(* CODESYS project PLC Pool Water Level Control Program.export

Project tree, tasks and I/O mapping:
  Device : CODESYS Control Win V3 x64, CODESYS, version 3.5.22.40
    application Application
      libraries: Standard, 3.5.22.0 (System)
      task MainTask (cyclic, interval t#100ms, priority 1) calls PLC_PRG [Read level and calculate pump command], TankSimulation [Use the command to calculate the new tank volume], TrialTester, TuningManager
      task VISU_TASK (cyclic, interval 100 ms, priority 31) calls VisuElems.Visu_Prg
      program PLC_PRG [LD]
      function block PoolModel [ST]
      program TankSimulation [ST]
      program TrialTester [ST]
      program TuningManager [ST]
      function block TuningTrial [ST]
      function block Twiddle [ST]
      function block ValveController [ST]
      visualisation TankOverview
*)

// Device/Application/PLC_PRG
PROGRAM PLC_PRG
VAR
	AutomationEnabled: BOOL; // FALSE means system is in manual mode
	ValveCommand : REAL := 0.0; // this is the precent-open that the valve needs to be
	FillingRequest : BOOL := FALSE;
	LowLevel : BOOL := FALSE; // when tank reaches 30% or less
	HighLevel : BOOL := FALSE; // when tank reaches 80% or more
	Trip : BOOL := FALSE; // activated automatically when HighHigh becomes TRUE
	ResetTrip : BOOL := FALSE;  // activated by operator switch
	
	// configure the controller
	LevelController : ValveController;
END_VAR

VAR_INPUT
	PoolLevelDeviation : REAL := 0.0; // inches
	HighHigh : BOOL := FALSE; // when level reaches 95% due to a system errors
	ActiveKp : REAL := 40.0;
	ActiveKi : REAL := 1.0;
END_VAR

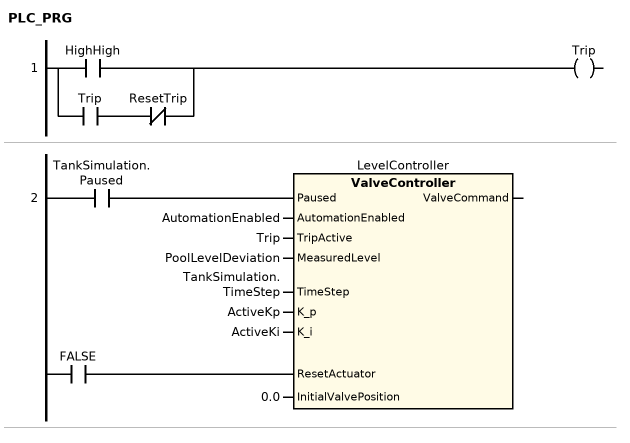
// NETWORK 1
Trip := HighHigh OR Trip AND NOT ResetTrip;

// NETWORK 2
LevelController(
    Paused := TankSimulation.Paused,
    AutomationEnabled := AutomationEnabled,
    TripActive := Trip,
    MeasuredLevel := PoolLevelDeviation,
    TimeStep := TankSimulation.TimeStep,
    K_p := ActiveKp,
    K_i := ActiveKi,
    ResetActuator := FALSE,
    InitialValvePosition := 0.0); // ValveController

END_PROGRAM

// Device/Application/ValveController
FUNCTION_BLOCK ValveController
VAR_INPUT
	Paused : BOOL;
	AutomationEnabled : BOOL := FALSE;
	TripActive : BOOL := FALSE;
	MeasuredLevel : REAL := 0.0; // inches. Positive means it's above the nomial level
	TimeStep : REAL := 0.1; //seconds 
	K_p : REAL := 1.0; // proportional tuning constant
	K_i : REAL := 1.0; // integral tuning contsant
	
	// to model a gradual response rather than instantaneous
	ResetActuator : BOOL := FALSE;
	InitialValvePosition : REAL := 0.0;
END_VAR
VAR_OUTPUT
	ValveCommand : REAL := 0.0; // percent to open
END_VAR
VAR
	// controller variables
	e : REAL := 0.0; // error
	P : REAL := 0.0; // proportional component
	I : REAL := 0.0; // integral component	
	u : REAL := 0.0; // valve command placeholder
	
	// for gradual response
	TargetValveCommand : REAL;
	MaxMove : REAL;
	ValveTravelTime : REAL := 20.0; // seconds to go from fully closed to fully open or vice versa 
	PreviousKp : REAL;
	PreviousKi : REAL;
	HasPreviousGains : BOOL := FALSE;
END_VAR

IF ResetActuator THEN
	ValveCommand := MAX(0.0, MIN(100.0, InitialValvePosition));
	TargetValveCommand := ValveCommand;
	I := 0.0;
	
	PreviousKp := K_p;
	PreviousKi := K_i;
	HasPreviousGains := TRUE;
	RETURN;
END_IF;

IF Paused THEN
	RETURN;
END_IF;

IF AutomationEnabled AND NOT TripActive THEN
	e := - MeasuredLevel;
	P := K_p * e;
	
	// match the new controller output to the current valve position
	IF HasPreviousGains AND ((K_p <> PreviousKp) OR (K_i <> PreviousKi)) THEN
		I := ValveCommand - P;
	END_IF;
	
	I := I + K_i * e * TimeStep;
	u := P + I;
	
	// prevent integral windup
	IF ((u > 100.0) AND (e > 0.0)) OR ((u < 0.0) AND (e < 0.0)) THEN
		I := I - K_i * e * TimeStep; // restore previous value
	END_IF;
	
	TargetValveCommand := MAX(0.0, MIN(100.0, P + I));
	
ELSE
	TargetValveCommand := 0.0;
	I := 0.0; // reset I
END_IF;

// Move actual valve position towards controller output
MaxMove := (100.0 / ValveTravelTime) * TimeStep;

ValveCommand := ValveCommand + MAX(-MaxMove, MIN(MaxMove, TargetValveCommand - ValveCommand));

ValveCommand := MAX(0.0, MIN(100.0, ValveCommand));

PreviousKp := K_p;
PreviousKi := K_i;
HasPreviousGains := TRUE;

END_FUNCTION_BLOCK

// Device/Application/TankSimulation
PROGRAM TankSimulation
VAR
	// pool data
	Volume : REAL := 100000.0; // current pool volume gal
	NominalVolume : REAL := 100000.0; // volume at target WL in gal
	SurfaceArea : REAL := 2500.0; // sq ft
	
	// physical constants
	MaxFillFlow : REAL := 50; // gpm, typical for 2" fill line
	EvapPerDay : REAL := 2; // inches
	SplashPerBather : REAL := 5.0; // splash loss (gal per hr)
	RainPerHour : REAL := 2.0; // inches
	LeakRate : REAL := 15.0; // gpm
	BackwashDuration : REAL := 300.0; // five minutes
	BackWashRate : REAL := 150.0; // gpm
	
	// inputs
	BatherCount : INT := 0; // current occupancy
	StartBackwash : BOOL := FALSE;
	StopBackwash : BOOL := FALSE;
	
	// Status variables
	PoolType : STRING := 'Outdoor'; // other option is 'Indoor'
	RainEnabled : BOOL := FALSE;
	LeakEnabled : BOOL := FALSE; 
	BackwashActive : BOOL := FALSE;
	BackwashElapsed : REAL := 0.0; // seconds
	SensorFailed: BOOL := FALSE;
	
	// Calculated values
	FillFlow: REAL := 0.0; // gpm
	EvapFlow : REAL := 0.0; // gpm
	SplashFlow : REAL := 0.0; // gpm
	RainFlow : REAL := 0.0; // gpm
	LeakFlow: REAL := 0.0; // gpm
	BackWashFlow : REAL := 0.0; // gpm
	WaterLevelDeviation: REAL := 0.0; // inches
	
	// time values
	TimeStep : REAL := 0.1; // s
	Paused : BOOL := FALSE; // user pauses the simulation to re-calibrate
	SensorLag : REAL := 5.0;
	MeasuredLevel : REAL := 0.0;
END_VAR

IF NOT Paused THEN
	IF PoolType = 'Indoor' THEN
		EvapFlow := (SurfaceArea / 12) * 7.48052 * (EvapPerDay / 1440);
	ELSIF PoolType = 'Outdoor' THEN
		EvapFlow := (SurfaceArea / 12) * 7.48052 * (EvapPerDay * 2 / 1440);
	ELSE
		EvapFlow := 0;
	END_IF;
	
	SplashFlow := BatherCount * SplashPerBather / 60;
	
	IF RainEnabled THEN
		RainFlow := (SurfaceArea * 7.48052 / (12 * 60)) * RainPerHour;
	ELSE
		RainFlow := 0;
	END_IF;
	
	
	IF LeakEnabled THEN
		LeakFlow := LeakRate; 
	ELSE
		LeakFlow := 0;
	END_IF;
	
	
	IF StartBackwash AND NOT StopBackwash THEN
		BackwashActive := TRUE;
	END_IF;
	
	IF StopBackwash THEN
		BackwashActive := FALSE;
		BackwashElapsed := 0.0;
	END_IF;
	
	IF BackwashElapsed >= BackwashDuration THEN
		BackwashActive := FALSE;
		BackwashElapsed := 0.0;
	END_IF;
	
	IF BackWashActive THEN
		BackwashFlow := BackwashRate;
		BackwashElapsed := BackwashElapsed + TimeStep;
	ELSE
		BackwashFlow := 0;
	END_IF;
	
	
	FillFlow := MaxFillFlow * (PLC_PRG.LevelController.ValveCommand / 100);
	
	// update volume
	Volume := Volume + (FillFlow + RainFlow - EvapFlow - SplashFlow - LeakFlow - BackwashFlow) * TimeStep / 60;
	WaterLevelDeviation := 12.0 * ((Volume - NominalVolume) / 7.48052) / SurfaceArea;
	
	// Simulate a failed sensor condition where it is stuck at a below-nominal reading
	IF SensorFailed THEN
		MeasuredLevel := -1.0; 
	ELSE
		MeasuredLevel := MeasuredLevel + (1.0 - EXP(-TimeStep / SensorLag)) * (WaterLevelDeviation - MeasuredLevel);
	END_IF;
	
	PLC_PRG.PoolLevelDeviation := MeasuredLevel;
	
	PLC_PRG.HighHigh := WaterLevelDeviation >= 1.0; // calculated independently of PoolLevel to be safe from sensor malfunctions
	
END_IF;

END_PROGRAM

// Device/Application/TrialTester
PROGRAM TrialTester
VAR
	TestTrial : TuningTrial;
	StartTest : BOOL := FALSE;
END_VAR

TestTrial(
	Start       := StartTest,
	CandidateKp := 40.0,
	CandidateKi := 1.0,
	InitialVolume := 99610.4, // includes an initial disturbance from the norm
	InitialMeasuredLevel := -0.25,
	TimeStep := 0.1,
	TrialDuration := 100.0,
	PoolType := 'Indoor',
	BatherCount := 0,
	MaxFillFlow := 50.0,
	EvapPerDay := 0.0,
	SplashPerBather := 0.0,
	RainPerHour := 0.0,
	LeakRate := 0.0,
	RainEnabled := FALSE,
	LeakEnabled := FALSE,
	SensorLag := 0.0
	);
	
StartTest := FALSE;

END_PROGRAM

// Device/Application/TuningTrial
FUNCTION_BLOCK TuningTrial
VAR_INPUT
	Start : BOOL; // to initialize trial
	CandidateKp : REAL;
	CandidateKi : REAL;
	InitialVolume : REAL;
	InitialMeasuredLevel : REAL;
	InitialValvePosition : REAL;
	TimeStep : REAL;
	TrialDuration : REAL; // length of simulation to run
	
	// to be imported from PoolModel
	PoolType          : STRING; // 'Indoor' or 'Outdoor' 
	BatherCount   : INT := 0; // current occupancy
	MaxFillFlow       : REAL := 50.0; // gpm, typical for 2" fill line
	EvapPerDay        : REAL; // inches - scale x2 for outdoor
	SplashPerBather   : REAL; // splash loss (gal per hr)
	RainPerHour       : REAL; // inches
	LeakRate          : REAL; // gpm
	RainEnabled       : BOOL := FALSE;
	LeakEnabled       : BOOL := FALSE; 
	SensorLag          : REAL; // s
END_VAR
VAR_OUTPUT
	Busy : BOOL; // whether trial is running
	Done : BOOL;
	Score : LREAL; // cumulative trial score
	Failed : BOOL := FALSE; // invalid or high-tripped trial
END_VAR
VAR
	TrialPool : PoolModel; // simulation model used for testing gain parameters
	TrialController : ValveController; 
	StepDuration : REAL;
	Elapsed : REAL; // s
END_VAR

IF Start THEN
	// reset Failed parameter
	Failed := FALSE;
	Score := 0.0;
	Elapsed := 0.0;
	
	// validate time parameters
	IF TimeStep <= 0.0 OR TrialDuration <= 0.0 THEN
		Busy := FALSE;
		Done := TRUE;
		Failed := TRUE;
	ELSE
		Score := 0.0;
		Elapsed := 0.0;
		TrialPool(
			Reset := TRUE,
			InitialVolume := InitialVolume,
			InitialMeasuredLevel := InitialMeasuredLevel,
			PoolType := PoolType,
			TimeStep := TimeStep,
			SensorLag := SensorLag,
			MaxFillFlow := MaxFillFlow,
			EvapPerDay := EvapPerDay,
			SplashPerBather := SplashPerBather,
			BatherCount := BatherCount,
			RainPerHour := RainPerHour,
			RainEnabled := RainEnabled,
			LeakRate := LeakRate,
			LeakEnabled := LeakEnabled,
			ValveCommand := 0.0,
			StartBackwash := FALSE,
			StopBackwash := FALSE,
			SensorFailed := FALSE
			);
		
		TrialController(
				Paused := FALSE,
				AutomationEnabled := FALSE,
				TripActive := FALSE,
				MeasuredLevel := TrialPool.MeasuredLevel,
				TimeStep := TimeStep,
				K_p := CandidateKp,
				K_i := CandidateKi,
				ResetActuator := TRUE,
				InitialValvePosition := InitialValvePosition
				);
				
		Busy := TRUE;
		DONE := FALSE;
	END_IF;
	
		
ELSIF Busy THEN
	IF TrialPool.HighHigh THEN
		Busy := FALSE;
		Done := TRUE;
		Failed := TRUE;
	ELSE
		StepDuration := MAX(0.0, MIN(TimeStep, TrialDuration - Elapsed));
		
		TrialController(
			Paused := FALSE,
			AutomationEnabled := TRUE,
			TripActive := FALSE,
			MeasuredLevel := TrialPool.MeasuredLevel,
			TimeStep := StepDuration,
			K_p := CandidateKp,
			K_i := CandidateKi,
			ResetActuator := FALSE
		);
		
		TrialPool(
			Reset := FALSE,
			InitialVolume := InitialVolume,
			InitialMeasuredLevel := InitialMeasuredLevel,
			PoolType := PoolType,
			TimeStep := StepDuration,
			SensorLag := SensorLag,
			MaxFillFlow := MaxFillFlow,
			EvapPerDay := EvapPerDay,
			SplashPerBather := SplashPerBather,
			BatherCount := BatherCount,
			RainPerHour := RainPerHour,
			RainEnabled := RainEnabled,
			LeakRate := LeakRate,
			LeakEnabled := LeakEnabled,
			ValveCommand := TrialController.ValveCommand,
			StartBackwash := FALSE,
			StopBackwash := FALSE,
			SensorFailed := FALSE
		);
		
		// check high limit again in case duration has been reached
		IF TrialPool.HighHigh THEN
			Busy := FALSE;
			Done := TRUE;
			Failed := TRUE;
		END_IF;
		
		Score := Score + ABS(TrialPool.ActualLevel) * StepDuration;
		Elapsed := Elapsed + StepDuration;
	
	END_IF;
	
	IF Elapsed >= TrialDuration THEN
		Busy := FALSE;
		Done := TRUE;
	END_IF;
	
END_IF;

END_FUNCTION_BLOCK

// Device/Application/PoolModel
FUNCTION_BLOCK PoolModel
VAR_INPUT
	
	// pool metrics
	PoolType           : STRING; // 'Indoor' or 'Outdoor' 
	InitialVolume      : REAL := 100000;   // wherever pool was at when auto tuning started
	
	// data
	Reset              : BOOL; // return to initial conditions
	InitialMeasuredLevel : REAL; // inches (from stilling well)
	ValveCommand       : REAL; // %
	TimeStep           : REAL; // s
	SensorLag          : REAL; // s
	
	// physical constants
	MaxFillFlow       : REAL := 50.0; // gpm, typical for 2" fill line
	EvapPerDay        : REAL; // inches - scale x2 for outdoor
	SplashPerBather   : REAL; // splash loss (gal per hr)
	RainPerHour       : REAL; // inches
	LeakRate          : REAL; // gpm
	BackwashDuration  : REAL := 300.0; // five minutes
	BackWashRate      : REAL := 150.0; // gpm
	
	// inputs
	BatherCount   : INT := 0; // current occupancy
	StartBackwash : BOOL := FALSE;
	StopBackwash  : BOOL := FALSE;
	
	// Status variables
	RainEnabled  : BOOL := FALSE;
	LeakEnabled  : BOOL := FALSE; 
	SensorFailed : BOOL := FALSE;
	
END_VAR
VAR_OUTPUT
	Volume        : REAL; // current volume in gal
	ActualLevel   : REAL; // inches
	MeasuredLevel : REAL; // inches (from sensor)
	FillFlow      : REAL; // gpm
	HighHigh      : BOOL; 
END_VAR
VAR
	CorrectedValveCommand : REAL := 0.0; // % 0 <= x <= 100
	SensorLevel         : REAL;	
	NominalVolume       : REAL := 100000.0; // gal
	SurfaceArea         : REAL := 2500.0; // sq ft
	EvapFlow            : REAL := 0.0; // gpm
	SplashFlow          : REAL := 0.0; // gpm
	RainFlow            : REAL := 0.0; // gpm
	LeakFlow            : REAL := 0.0; // gpm
	BackwashFlow        : REAL := 0.0; // gpm
	BackwashActive      : BOOL := FALSE;
	BackwashElapsed     : REAL := 0.0; // seconds
	BackwashTimeStep    : REAL := 0.0; // s
END_VAR

IF Reset THEN
	Volume := InitialVolume;
	BackwashActive := FALSE;
	BackwashElapsed := 0.0;
	BackwashFlow := 0.0;
	FillFlow := 0.0;
	EvapFlow := 0.0; // gpm
	SplashFlow := 0.0; // gpm
	RainFlow := 0.0; // gpm
	LeakFlow := 0.0;
ELSE
	IF PoolType = 'Indoor' THEN
		EvapFlow := (SurfaceArea / 12) * 7.48052 * (EvapPerDay / 1440);
	ELSIF PoolType = 'Outdoor' THEN
		EvapFlow := (SurfaceArea / 12) * 7.48052 * (EvapPerDay * 2 / 1440);
	ELSE
		EvapFlow := 0;
	END_IF;
	
	SplashFlow := BatherCount * SplashPerBather / 60;
	
	IF RainEnabled THEN
		RainFlow := (SurfaceArea * 7.48052 / (12 * 60)) * RainPerHour;
	ELSE
		RainFlow := 0;
	END_IF;
	
	
	IF LeakEnabled THEN
		LeakFlow := LeakRate; 
	ELSE
		LeakFlow := 0;
	END_IF;
	
	// use time remaining for backwash if it is less than TimeStep
	BackwashTimeStep := MAX(0.0, MIN(TimeStep, BackwashDuration - BackwashElapsed));
	
	IF StartBackwash AND NOT StopBackwash THEN
		BackwashActive := TRUE;
	END_IF;
	
	IF StopBackwash THEN
		BackwashActive := FALSE;
		BackwashElapsed := 0.0;
	END_IF;
	
	IF BackwashElapsed >= BackwashDuration THEN
		BackwashActive := FALSE;
		BackwashElapsed := 0.0;
	END_IF;
	
	IF BackWashActive THEN
		BackwashFlow := BackwashRate;
		BackwashElapsed := BackwashElapsed + BackwashTimeStep;
	ELSE
		BackwashFlow := 0;
	END_IF;

	
	IF ValveCommand > 100 THEN
		CorrectedValveCommand := 100;
	ELSIF ValveCommand < 0 THEN
		CorrectedValveCommand := 0;
	ELSE
		CorrectedValveCommand := ValveCommand;
	END_IF;
	FillFlow := MaxFillFlow * (CorrectedValveCommand / 100);
	
	// update volume
	Volume := Volume + (FillFlow + RainFlow - EvapFlow - SplashFlow - LeakFlow) * TimeStep / 60 - BackwashFlow * BackwashTimeStep / 60;
	
END_IF;
	
ActualLevel := 12.0 * ((Volume - NominalVolume) / 7.48052) / SurfaceArea;

// Simulate a failed sensor condition where it is stuck at a below-nominal reading
IF Reset THEN
	MeasuredLevel := InitialMeasuredLevel;
ELSIF SensorFailed THEN
	MeasuredLevel := -1.0; 
ELSIF SensorLag <= 0 THEN
	MeasuredLevel := ActualLevel;
ELSE
	MeasuredLevel := MeasuredLevel + (1 - EXP(-TimeStep / SensorLag)) * (ActualLevel - MeasuredLevel);
END_IF;

HighHigh := ActualLevel >= 1; // calculated independently of MeasuredLevel to be safe from sensor malfunctions

END_FUNCTION_BLOCK

// Device/Application/TuningManager
PROGRAM TuningManager
VAR
	Tuner : Twiddle;
	StartTuning : BOOL := FALSE; // pulse true to start tuning
END_VAR


Tuner(
	Start := StartTuning,
	InitialKp := PLC_PRG.ActiveKp,
	InitialKi := PLC_PRG.ActiveKi,
	InitialValvePosition := PLC_PRG.LevelController.ValveCommand,
	InitialVolume := TankSimulation.Volume,
	InitialMeasuredLevel := PLC_PRG.PoolLevelDeviation,
	PoolType := TankSimulation.PoolType,
	BatherCount := TankSimulation.BatherCount,
	MaxFillFlow := TankSimulation.MaxFillFlow,
	EvapPerDay := TankSimulation.EvapPerDay,
	SplashPerBather := TankSimulation.SplashPerBather,
	RainPerHour := TankSimulation.RainPerHour,
	LeakRate := TankSimulation.LeakRate,
	RainEnabled := TankSimulation.RainEnabled,
	LeakEnabled := TankSimulation.LeakEnabled,
	SensorLag := 5.0 // seconds
	);
	
IF Tuner.Done AND Tuner.HasValidBest AND NOT Tuner.Failed THEN
	PLC_PRG.ActiveKp := Tuner.BestKp;
	PLC_PRG.ActiveKi := Tuner.BestKi;
END_IF;

StartTuning := FALSE;

END_PROGRAM

// Device/Application/Twiddle
FUNCTION_BLOCK Twiddle
VAR_INPUT
	Start : BOOL; // one-call pulse to begin tuning
	InitialKp : REAL;
	InitialKi : REAL;
	InitialValvePosition : REAL;
	
	// pool data
	InitialVolume : REAL;
	InitialMeasuredLevel : REAL;
	
	// environmental settings
	PoolType          : STRING; // 'Indoor' or 'Outdoor' 
	BatherCount   : INT := 0; // current occupancy
	MaxFillFlow       : REAL := 50.0; // gpm, typical for 2" fill line
	EvapPerDay        : REAL; // inches - scale x2 for outdoor
	SplashPerBather   : REAL; // splash loss (gal per hr)
	RainPerHour       : REAL; // inches
	LeakRate          : REAL; // gpm
	RainEnabled       : BOOL := FALSE;
	LeakEnabled       : BOOL := FALSE; 
	SensorLag          : REAL; // s
END_VAR

VAR_OUTPUT
	Busy : BOOL;
	Done : BOOL;
	Failed : BOOL;
	Converged : BOOL; // if optimization thresholds were reached
	
	BestKp : REAL; 
	BestKi : REAL;
	BestScore : LREAL;
	HasValidBest : BOOL; // whether any trial was successful
END_VAR

VAR
	// data parameters
	TimeStep : REAL := 0.1; // s
	TrialDuration : REAL := 100.0; // s
	Trial : TuningTrial; // evaluate candidate gains
	State : INT := 0; // current stage of the search
	StepIndex : INT;
	StepsPerScan : INT := 1000; // to speed up the computation
	
	// gain-related variables
	ParameterIndex : INT; // Which gain is being adjusted
	TestKp : REAL := 40.0; // Starting point
	TestKi : REAL := 1.0; // Starting point
	DeltaKp : REAL := 10.0; // search increments
	DeltaKi : REAL := 0.25;                                                                                                         
	Iteration : INT := 0; 
	TestingNegative : BOOL := FALSE; // whether a negative DeltaGain is being tested
	
	// snapshot variables to ignore conditions changing mid-tuning
	SnapshotVolume            : REAL;
	SnapshotMeasuredLevel     : REAL;
	SnapshotValvePosition     : REAL;
	SnapshotPoolType          : STRING; // 'Indoor' or 'Outdoor' 
	SnapshotBatherCount       : INT := 0; // current occupancy
	SnapshotMaxFillFlow       : REAL := 50.0; // gpm, typical for 2" fill line
	SnapshotEvapPerDay        : REAL; // inches - scale x2 for outdoor
	SnapshotSplashPerBather   : REAL; // splash loss (gal per hr)
	SnapshotRainPerHour       : REAL; // inches
	SnapshotLeakRate          : REAL; // gpm
	SnapshotRainEnabled       : BOOL := FALSE;
	SnapshotLeakEnabled       : BOOL := FALSE; 
	SnapshotSensorLag         : REAL; // s
	
	// optimization thresholds
	ToleranceKp : REAL := 0.1;
	ToleranceKi : REAL := 0.005;
	MaxIterations : INT := 100;
END_VAR

IF Start AND NOT Busy THEN
	Busy := TRUE;
	Done := FALSE;
	Failed := FALSE;
	Converged := FALSE;
	TestingNegative := FALSE;
	HasValidBest := FALSE;
	BestScore := 0.0;
	Iteration := 0;
	DeltaKp := 10.0;
	DeltaKi := 0.25;
	
	// initialize the stored gains
	BestKp := InitialKp;
	BestKi := InitialKi;
	TestKp := InitialKp;
	TestKi := InitialKi;
	
	// capture snapshot 
	SnapshotVolume          := InitialVolume;
	SnapshotMeasuredLevel   := InitialMeasuredLevel;
	SnapshotValvePosition   := InitialValvePosition;
	SnapshotPoolType        := PoolType;
	SnapshotBatherCount     := BatherCount;
	SnapshotMaxFillFlow     := MaxFillFlow;
	SnapshotEvapPerDay      := EvapPerDay;
	SnapshotSplashPerBather := SplashPerBather;
	SnapshotRainPerHour     := RainPerHour;
	SnapshotLeakRate        := LeakRate;
	SnapshotRainEnabled     := RainEnabled;
	SnapshotLeakEnabled     := LeakEnabled; 
	SnapshotSensorLag       := SensorLag;
	
	// advance to next stage
	State := 10;
END_IF;

CASE State OF
	0:
		// nothing
	
	10: 
		Trial(
			Start := TRUE,
			CandidateKp := TestKp,
			CandidateKi := TestKi,
			InitialVolume := SnapshotVolume,
			InitialMeasuredLevel := SnapshotMeasuredLevel,
			InitialValvePosition := SnapshotValvePosition,
			TimeStep := TimeStep,
			TrialDuration := TrialDuration,
			PoolType := SnapshotPoolType,
			BatherCount := SnapshotBatherCount,
			MaxFillFlow := SnapshotMaxFillFlow,
			EvapPerDay := SnapshotEvapPerDay,
			SplashPerBather := SnapshotSplashPerBather,
			RainPerHour := SnapshotRainPerHour,
			LeakRate := SnapshotLeakRate,
			RainEnabled := SnapshotRainEnabled,
			LeakEnabled := SnapshotLeakEnabled,			
			SensorLag := SnapshotSensorLag
			);
		
		State := 20;
	
	20:
		FOR StepIndex := 1 TO StepsPerScan DO
			Trial(
				Start := FALSE,
				CandidateKp := TestKp,
				CandidateKi := TestKi,
				InitialVolume := SnapshotVolume,
				InitialMeasuredLevel := SnapshotMeasuredLevel,
				InitialValvePosition := SnapshotValvePosition,
				TimeStep := TimeStep,
				TrialDuration := TrialDuration,
				PoolType := SnapshotPoolType,
				BatherCount := SnapshotBatherCount,
				MaxFillFlow := SnapshotMaxFillFlow,
				EvapPerDay := SnapshotEvapPerDay,
				SplashPerBather := SnapshotSplashPerBather,
				RainPerHour := SnapshotRainPerHour,
				LeakRate := SnapshotLeakRate,
				RainEnabled := SnapshotRainEnabled,
				LeakEnabled := SnapshotLeakEnabled,			
				SensorLag := SnapshotSensorLag
				);
				IF Trial.Done THEN
					EXIT;
				END_IF;
			END_FOR;
			
		IF Trial.Done THEN
			State := 30;
		END_IF;
	
	30:
		IF NOT Trial.Failed THEN
			BestScore := Trial.Score;
			HasValidBest := TRUE;
			
			// get ready to run Kp trial
			ParameterIndex := 0;
			TestKp := BestKp + DeltaKp;
			TestKi := BestKi;
			
			State := 40;
		ELSE
			Failed := TRUE;
			Busy := FALSE;
			Done := TRUE;
			State := 0; // end the search
		END_IF;
		
	40:
		Trial(
			Start := TRUE,
			CandidateKp := TestKp,
			CandidateKi := TestKi,
			InitialVolume := SnapshotVolume,
			InitialMeasuredLevel := SnapshotMeasuredLevel,
			InitialValvePosition := SnapshotValvePosition,
			TimeStep := TimeStep,
			TrialDuration := TrialDuration,
			PoolType := SnapshotPoolType,
			BatherCount := SnapshotBatherCount,
			MaxFillFlow := SnapshotMaxFillFlow,
			EvapPerDay := SnapshotEvapPerDay,
			SplashPerBather := SnapshotSplashPerBather,
			RainPerHour := SnapshotRainPerHour,
			LeakRate := SnapshotLeakRate,
			RainEnabled := SnapshotRainEnabled,
			LeakEnabled := SnapshotLeakEnabled,			
			SensorLag := SnapshotSensorLag
			);
			
		State := 50;
	
	50:
		FOR StepIndex := 1 TO StepsPerScan DO
			Trial(
				Start := FALSE,
				CandidateKp := TestKp,
				CandidateKi := TestKi,
				InitialVolume := SnapshotVolume,
				InitialMeasuredLevel := SnapshotMeasuredLevel,
				InitialValvePosition := SnapshotValvePosition,
				TimeStep := TimeStep,
				TrialDuration := TrialDuration,
				PoolType := SnapshotPoolType,
				BatherCount := SnapshotBatherCount,
				MaxFillFlow := SnapshotMaxFillFlow,
				EvapPerDay := SnapshotEvapPerDay,
				SplashPerBather := SnapshotSplashPerBather,
				RainPerHour := SnapshotRainPerHour,
				LeakRate := SnapshotLeakRate,
				RainEnabled := SnapshotRainEnabled,
				LeakEnabled := SnapshotLeakEnabled,			
				SensorLag := SnapshotSensorLag
				);
				IF Trial.Done THEN
					EXIT;
				END_IF;
			END_FOR;
		
		IF Trial.Done THEN
			State := 60;
		END_IF;
			
	60:
		
		IF NOT Trial.Failed AND Trial.Score < BestScore THEN
			BestScore := Trial.Score;
			BestKp := TestKp;
			BestKi := TestKi;
			IF ParameterIndex = 0 THEN
				DeltaKp := DeltaKp * 1.1;
			ELSIF ParameterIndex = 1 THEN
				DeltaKi := DeltaKi * 1.1;
			END_IF;
			State := 70; // to switch to the next parameter
		ELSE
			IF TestingNegative THEN
				// if positive and negative increments didn't improve the score then shrink the increment and move to the next gain
				IF ParameterIndex = 0 THEN
					DeltaKp := DeltaKp * 0.9; // shrink
				ELSIF ParameterIndex = 1 THEN
					DeltaKi := DeltaKi * 0.9; // shrink
				END_IF;
				State := 70; 
			ELSE
				// if positive increment didn't work then try a negative increment on the same gain parameter
				TestKp := BestKp;
				TestKi := BestKi;
				IF ParameterIndex = 0 THEN
					TestKp := MAX(0.0, BestKp - DeltaKp);
				ELSIF ParameterIndex = 1 THEN
					TestKi := MAX(0.0, BestKi - DeltaKi);
				END_IF;
				TestingNegative := TRUE;
				State := 40;
			END_IF;
		END_IF;
	
	70:
		IF ParameterIndex = 0 THEN
			ParameterIndex := 1;
		ELSIF ParameterIndex = 1 THEN
			ParameterIndex := 0;
			Iteration := Iteration + 1;
		END_IF;
		
		IF ((DeltaKp <= ToleranceKp) AND (DeltaKi <= ToleranceKi)) OR (Iteration >= MaxIterations) THEN
			Busy := FALSE;
			Done := TRUE;
			State := 0;
			Converged := (DeltaKp <= ToleranceKp) AND (DeltaKi <= ToleranceKi);
		ELSE
			TestingNegative := FALSE;
			TestKp := BestKp;
			TestKi := BestKi;
			IF ParameterIndex = 0 THEN
				TestKp := BestKp + DeltaKp;
			ELSIF ParameterIndex = 1 THEN
				TestKi := BestKi + DeltaKi;
			END_IF;
			State := 40;
		END_IF;
			
		
	
	
END_CASE;

END_FUNCTION_BLOCK

// Device/Application/TankOverview
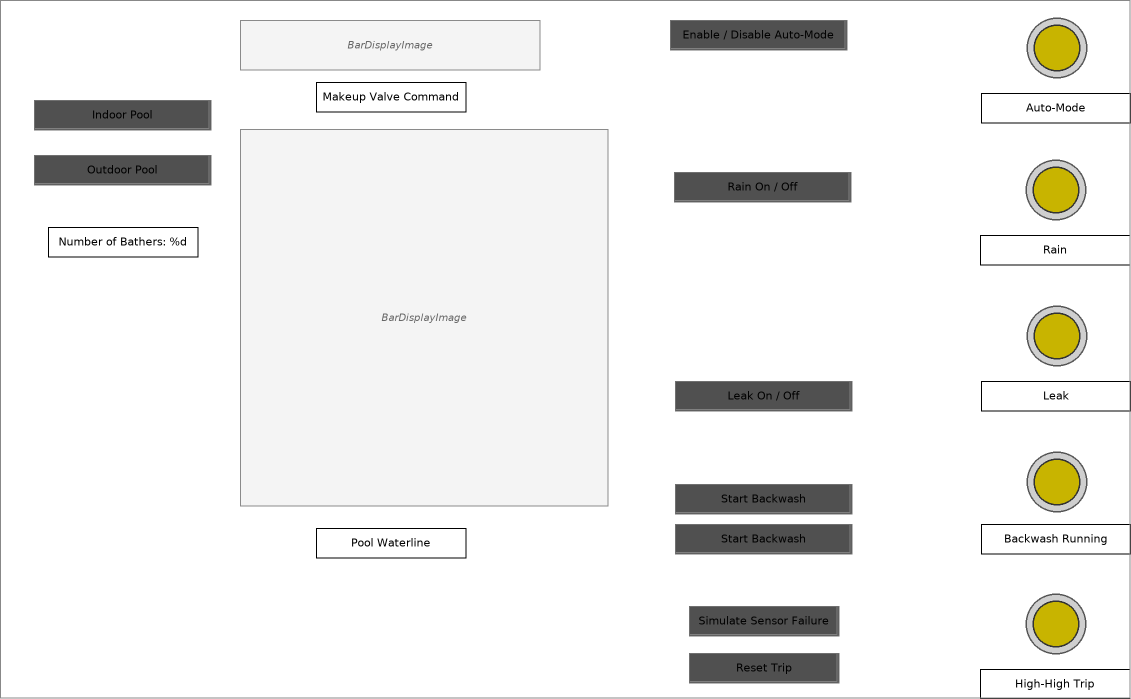
VISUALIZATION TankOverview  // 1131x699
    BarDisplayImage (240,129 368x377), value: TankSimulation.WaterLevelDeviation, style: BarDisplayImage-Gray, scale format: %.1f, scale -3..3
        p518627256: Inches
    Button (670,20 177x30), "Enable / Disable Auto-Mode"
        toggle PLC_PRG.AutomationEnabled
    Rectangle (316,82 150x30), "Makeup Valve Command"
    Lamp1 (1021,589 70x70), variable: PLC_PRG.Trip, style: Lamp-Lamp1-Yellow
    Rectangle (980,669 150x30), "High-High Trip"
    Button (689,653 150x30), "Reset Trip"
        tap PLC_PRG.ResetTrip
    Button (689,606 150x30), "Simulate Sensor Failure"
        toggle TankSimulation.SensorFailed
    BarDisplayImage (240,20 300x50), value: PLC_PRG.LevelController.ValveCommand, style: BarDisplayImage-Gray, scale format: %.1f, scale 0..100
        p518627256: %
    Rectangle (316,528 150x30), "Pool Waterline"
    Button (674,172 177x30), "Rain On / Off"
        toggle TankSimulation.RainEnabled
    Button (675,381 177x30), "Leak On / Off"
        toggle TankSimulation.LeakEnabled
    Button (675,484 177x30), "Start Backwash"
        toggle TankSimulation.StartBackwash
    Button (675,524 177x30), "Start Backwash"
        toggle TankSimulation.StopBackwash
    Lamp1 (1022,447 70x70), variable: TankSimulation.BackwashActive, style: Lamp-Lamp1-Yellow
    Rectangle (981,524 150x30), "Backwash Running"
    Lamp1 (1022,301 70x70), variable: TankSimulation.LeakEnabled, style: Lamp-Lamp1-Yellow
    Rectangle (981,381 150x30), "Leak"
    Lamp1 (1021,155 70x70), variable: TankSimulation.RainEnabled, style: Lamp-Lamp1-Yellow
    Rectangle (980,235 150x30), "Rain"
    Lamp1 (1022,13 70x70), variable: PLC_PRG.AutomationEnabled, style: Lamp-Lamp1-Yellow
    Rectangle (981,93 150x30), "Auto-Mode"
    Button (34,155 177x30), "Outdoor Pool", colour toggle: TankSimulation.PoolType = 'Outdoor'
        OnMouseClick: execute { TankSimulation.PoolType := 'Outdoor'; }
    Button (34,100 177x30), "Indoor Pool", colour toggle: TankSimulation.PoolType = 'Indoor'
        OnMouseClick: execute { TankSimulation.PoolType := 'Indoor'; }
    Rectangle (48,227 150x30), "Number of Bathers: %d", text variable: TankSimulation.BatherCount
        OnMouseClick: write the text variable via Edit, min 0, max 200
END_VISUALIZATION
